(* IEC 61131-3 sources: codesys-framework/txt/application/WeVe Core (library)/30 Module/Hardware/FB_Hardware, 3 files *)

(* ---- LoadHardCodedSettings.method.st ---- *)
METHOD PROTECTED ABSTRACT LoadHardCodedSettings
VAR_INPUT
END_VAR

// --- BEGIN IMPLEMENTATION ---

(* ---- ProcessErrors.method.st ---- *)
METHOD PROTECTED ProcessErrors
VAR_INPUT
END_VAR

// --- BEGIN IMPLEMENTATION ---

;

(* ---- ProcessHardware.method.st ---- *)
METHOD PROTECTED ABSTRACT ProcessHardware
VAR_INPUT
END_VAR

// --- BEGIN IMPLEMENTATION ---
